(* PLC project Storage_Main, Beckhoff Automation GmbH TwinCAT PLC Control 3.5.13.21 *)
(* stored: creationDateTime 2026-11-24T10:08:08.1458531, modificationDateTime 2026-11-24T10:08:08.1488473 *)

PROGRAM SFC_Test
VAR_INPUT
    SFCReset : BOOL;
END_VAR
VAR
    nTest : INT;
END_VAR

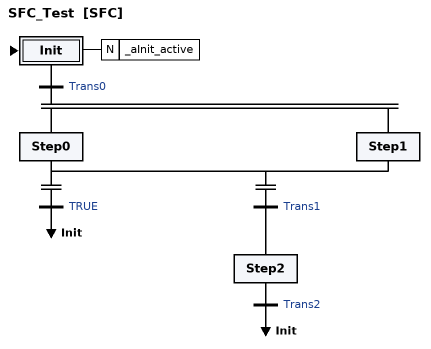
INITIAL_STEP Init:
  _aInit_active(N);
END_STEP
TRANSITION FROM Init TO (Step0, Step1)
  := Trans0;
END_TRANSITION
STEP Step0:
END_STEP
TRANSITION FROM (Step0, Step1) TO Init
  := TRUE;
END_TRANSITION
TRANSITION FROM (Step0, Step1) TO Step2
  := Trans1;
END_TRANSITION
STEP Step1:
END_STEP
STEP Step2:
END_STEP
TRANSITION FROM Step2 TO Init
  := Trans2;
END_TRANSITION

ACTION _aInit_active:
                
              
END_ACTION
END_PROGRAM
